Fanuc KAREL source: kb00043.KL

-- PROVISIONAL review KL for V770-1; original PC SHA256 999701eba7efd021aa1ee61e242c9dc2a6eab986fbf7d0f2214a2146d77c0016
-- Incomplete behavior may be omitted. Consult companion uncertainty JSON. Do not deploy.
PROGRAM KB00043
%NOLOCKGROUP
BEGIN
  -- UNRESOLVED_PC offsets 5-12; opcodes 9D,23
  -- UNRESOLVED_PC offsets 17-26; opcodes 3F,75
  -- UNRESOLVED_PC offsets 31-49; opcodes 27,22,22,2A,31
  -- UNRESOLVED_PC offsets 54-58; opcodes 7F
END KB00043
